(* IEC 61131-3 sources: Enumium/projects/downhome-spice-line/software/plc, 4 files *)

(* ---- DosingStation.st ---- *)
(* ============================================================================
   P1-225  PHASE 1 DOSING STATION  (IEC 61131-3 ST, CODESYS 3.5 on WAGO PFC200 750-8212)
   Down Home Creole Phase 1 prototype. Ring of up to 12 ingredient bins
   (P1-211) with 2 in volumetric screw feeders (P1-212, VFD P1-226) dosing
   one at a time into weigh hopper P1-220 (3 x 50 kg cells, Rice Lake 880
   indicator P1-222, 10 g division). When the list is done, butterfly valve
   P1-223 opens and flexible screw P1-224 carries the charge to blender P1-301
   (on riser stand P1-311). The hand-weighed lines and the premix are then
   tipped into the screw's intake grate, so nobody lifts a pail above waist height.

   The MES owns the recipe and the lot genealogy:
     GET /api/batch/<id>/doselist  -> MES_DoseList (largest dose first)
     POST /api/dose {batch, bin, actual_kg} after each finished dose.
   The PLC owns the equipment: one feeder at a time, never a screw into a
   closed valve or a full blender, no dose from a bin at low level.

   Dosing method (gain in weight, per bin):
     FAST  : VFD at FastHz until  net >= target - SlowBand - InFlight
     SLOW  : VFD at SlowHz until  net >= target - InFlight
     SETTLE: feeder off, wait SettleT, read stable weight
     CHECK : |actual - target| <= TolKg  -> report;  under -> one JOG pulse
             (max 3) ;  over -> OVERDOSE alarm, hold for the operator.
   In-flight (material still falling after the screw stops) is learned per
   bin: InFlight := InFlight + 0.5 * (actual - target), clamped 0..0.5 kg.
   No-flow: hopper gain < 0.05 kg in NoFlowT while the feeder runs -> alarm
   (bridged bin, empty bin, broken shear pin).
   Timers and speeds marked (SAT) are tuned at site acceptance.
   E-stop and the hopper/screw guards are hard-wired through safety relay
   SR-P1 and remove VFD enable; this code only sees the healthy bit.
   ============================================================================ *)

TYPE E_DoseStep : (
    IDLE := 0, WAIT_LIST := 5, PRECHECK := 10, TARE := 20, FAST := 30, SLOW := 40,
    SETTLE := 50, CHECK := 60, JOG := 65, REPORT := 70, NEXT := 80,
    TRANSFER := 90, TRANSFER_DRAIN := 95, COMPLETE := 100, HELD := 110, ABORTED := 120 );
END_TYPE

TYPE ST_DoseStep :
STRUCT
    Bin        : INT;          (* 1..12, ring position *)
    Ingredient : STRING[24];
    TargetKg   : REAL;         (* >= 4 kg by MES rule *)
    TolKg      : REAL;         (* max(1 % of target, 0.02 kg) *)
END_STRUCT
END_TYPE

TYPE ST_DoseList :
STRUCT
    BatchID  : STRING[16];
    FormulaID: STRING[16];
    Steps    : ARRAY[1..12] OF ST_DoseStep;
    Count    : INT;
    Valid    : BOOL;
END_STRUCT
END_TYPE

TYPE ST_DoseResult :
STRUCT
    BatchID  : STRING[16];
    Bin      : INT;
    ActualKg : REAL;
    Ready    : BOOL;           (* MES gateway posts /api/dose then sets Ack *)
    Ack      : BOOL;
END_STRUCT
END_TYPE

VAR_GLOBAL CONSTANT
    NBINS        : INT  := 12;
    HOPPER_MAXKG : REAL := 100.0;   (* 3 x 50 kg cells, 2/3 derated for the hopper *)
    BLENDER_MAXKG: REAL := 95.0;    (* P1-301 6 cu ft x densest blend (0.56 g/ml) *)
END_VAR

VAR_GLOBAL
    (* ---- I/O (WAGO 750-8212 rack: 750-430 DI, 750-530 DO, 750-455 AI 4-20 mA, Modbus RTU to GS20 drives) ---- *)
    DI_SafetyOK      AT %IX0.0  : BOOL;     (* SR-P1 healthy: e-stops, hopper lid, screw guard *)
    DI_ValveClosed   AT %IX0.1  : BOOL;     (* P1-223 closed limit *)
    DI_ValveOpen     AT %IX0.2  : BOOL;     (* P1-223 open limit *)
    DI_ScrewRunning  AT %IX0.3  : BOOL;     (* P1-224 motor contactor aux *)
    DI_BlenderReady  AT %IX0.4  : BOOL;     (* P1-301 cover closed and not discharging *)
    DI_BlenderHigh   AT %IX0.5  : BOOL;     (* P1-301 high level, capacitance probe *)
    DI_DustFanOn     AT %IX0.6  : BOOL;     (* P1-310 fan running *)
    DI_BinLow        AT %IX1.0  : ARRAY[1..12] OF BOOL;   (* P1-213 Soliphant FTM20, TRUE = covered (fail-safe) *)
    DO_ValveOpen     AT %QX0.0  : BOOL;     (* P1-223 solenoid *)
    DO_ScrewRun      AT %QX0.1  : BOOL;     (* P1-224 contactor *)
    DO_Horn          AT %QX0.2  : BOOL;
    DO_Beacon        AT %QX0.3  : BOOL;
    DO_Agitator      AT %QX1.0  : ARRAY[1..12] OF BOOL;   (* bin flow aid, density < 0.5 kg/L bins only *)
    AI_HopperKg                 : REAL;     (* P1-222 Rice Lake 880 gross weight over Modbus TCP, 10 g *)
    AI_HopperStable             : BOOL;     (* 880 motion bit inverted *)
    VFD_Run          : ARRAY[1..12] OF BOOL;      (* GS20 drives, Modbus RTU *)
    VFD_Hz           : ARRAY[1..12] OF REAL;
    VFD_Fault        : ARRAY[1..12] OF BOOL;

    (* ---- MES interface (OPC UA server on the PFC200, written by the MES gateway) ---- *)
    MES_DoseList     : ST_DoseList;
    MES_Result       : ST_DoseResult;
    MES_Start        : BOOL;
    MES_HandAddsDone : BOOL;            (* hand-weighed lines, then the premix, tipped into the P1-224 intake grate *)
    MES_Abort        : BOOL;
    HMI_Resume       : BOOL;
    HMI_Reset        : BOOL;

    (* ---- status ---- *)
    Dose_Step        : E_DoseStep;
    Dose_Index       : INT;
    Dose_NetKg       : REAL;
    Dose_Alarm       : STRING[60];
    Dose_HeldFrom    : E_DoseStep;

    (* ---- per-bin parameters, retained (learned in-flight survives power loss) ---- *)
    InFlightKg       : ARRAY[1..12] OF REAL := [12(0.15)];   (* (SAT) start value *)
    FastHz           : ARRAY[1..12] OF REAL := [12(60.0)];   (* about 700 L/h at 60 Hz, 2 in screw *)
    SlowHz           : ARRAY[1..12] OF REAL := [12(12.0)];   (* (SAT) *)
    SlowBandKg       : ARRAY[1..12] OF REAL := [12(1.0)];    (* (SAT) *)
END_VAR

PROGRAM DosingStation
VAR
    tStep     : TON;
    tNoFlow   : TON;
    tSettle   : TON;
    tTransfer : TON;
    TareKg    : REAL;
    LastKg    : REAL;
    ActualKg  : REAL;
    Jogs      : INT;
    i         : INT;
    b         : INT;           (* bin of the current step *)
    s         : ST_DoseStep;
    SumKg     : REAL;
    NoFlowT   : TIME := T#8S;  (* (SAT) *)
    SettleT   : TIME := T#3S;  (* (SAT) *)
    JogT      : TIME := T#600MS;
    DrainT    : TIME := T#20S; (* screw runs on after the hopper reads empty *)
    MaxDoseT  : TIME := T#10M; (* longest planned dose < 8 min *)
END_VAR

(* ---------- always: interlocks ---------- *)
IF NOT DI_SafetyOK OR MES_Abort THEN
    FOR i := 1 TO NBINS DO VFD_Run[i] := FALSE; END_FOR
    DO_ScrewRun := FALSE;
    DO_ValveOpen := FALSE;
    IF Dose_Step <> IDLE AND Dose_Step <> COMPLETE THEN
        Dose_Alarm := SEL(MES_Abort, 'SAFETY CIRCUIT OPEN', 'ABORTED BY MES');
        Dose_Step := ABORTED;
    END_IF
END_IF

(* the transfer screw may only run with the valve open, the blender ready and the dust fan on *)
IF DO_ScrewRun AND NOT (DI_ValveOpen AND DI_BlenderReady AND DI_DustFanOn AND NOT DI_BlenderHigh) THEN
    DO_ScrewRun := FALSE;
    DO_ValveOpen := FALSE;
    Dose_Alarm := 'TRANSFER PERMISSIVE LOST';
    Dose_HeldFrom := Dose_Step;
    Dose_Step := HELD;
END_IF

(* one feeder at a time: only the current bin may run *)
FOR i := 1 TO NBINS DO
    IF VFD_Run[i] AND ((Dose_Step <> FAST AND Dose_Step <> SLOW AND Dose_Step <> JOG) OR i <> b) THEN
        VFD_Run[i] := FALSE;
    END_IF
    IF VFD_Fault[i] AND VFD_Run[i] THEN
        VFD_Run[i] := FALSE;
        Dose_Alarm := CONCAT('FEEDER FAULT BIN ', INT_TO_STRING(i));
        Dose_HeldFrom := Dose_Step;
        Dose_Step := HELD;
    END_IF
    DO_Agitator[i] := VFD_Run[i];       (* flow aid only while its feeder runs *)
END_FOR

Dose_NetKg := AI_HopperKg - TareKg;

(* ---------- sequence ---------- *)
CASE Dose_Step OF

IDLE:
    IF MES_Start THEN Dose_Step := WAIT_LIST; END_IF

WAIT_LIST:
    IF MES_DoseList.Valid AND MES_DoseList.Count >= 1 AND MES_DoseList.Count <= NBINS THEN
        SumKg := 0.0;
        FOR i := 1 TO MES_DoseList.Count DO SumKg := SumKg + MES_DoseList.Steps[i].TargetKg; END_FOR
        IF SumKg > HOPPER_MAXKG OR SumKg > BLENDER_MAXKG THEN
            Dose_Alarm := 'DOSE LIST EXCEEDS HOPPER OR BLENDER';
            Dose_Step := ABORTED;
        ELSE
            Dose_Index := 1;
            Dose_Step := PRECHECK;
        END_IF
    END_IF

PRECHECK:
    (* hopper empty, valve closed, dust fan on *)
    IF NOT DI_DustFanOn THEN
        Dose_Alarm := 'DUST COLLECTOR P1-310 OFF';
    ELSIF NOT DI_ValveClosed THEN
        Dose_Alarm := 'HOPPER VALVE NOT CLOSED';
    ELSIF AI_HopperKg > 0.5 THEN
        Dose_Alarm := 'HOPPER NOT EMPTY';
    ELSE
        Dose_Alarm := '';
        Dose_Step := TARE;
    END_IF

TARE:
    s := MES_DoseList.Steps[Dose_Index];
    b := s.Bin;
    IF b < 1 OR b > NBINS THEN
        Dose_Alarm := 'BAD BIN NUMBER IN DOSE LIST';
        Dose_Step := ABORTED;
    ELSIF NOT DI_BinLow[b] THEN
        Dose_Alarm := CONCAT('BIN LOW: REFILL BIN ', INT_TO_STRING(b));   (* MES checked book stock; this is the probe *)
        Dose_HeldFrom := TARE;
        Dose_Step := HELD;
    ELSIF AI_HopperStable THEN
        TareKg := AI_HopperKg;        (* cumulative: each dose is tared on the previous ones *)
        LastKg := AI_HopperKg;
        Jogs := 0;
        VFD_Hz[b] := FastHz[b];
        VFD_Run[b] := TRUE;
        Dose_Step := FAST;
    END_IF

FAST, SLOW:
    IF Dose_Step = FAST AND Dose_NetKg >= s.TargetKg - SlowBandKg[b] - InFlightKg[b] THEN
        VFD_Hz[b] := SlowHz[b];
        Dose_Step := SLOW;
    ELSIF Dose_NetKg >= s.TargetKg - InFlightKg[b] THEN
        VFD_Run[b] := FALSE;
        Dose_Step := SETTLE;
    END_IF
    (* no-flow: the hopper must gain 50 g in NoFlowT *)
    tNoFlow(IN := VFD_Run[b] AND (AI_HopperKg - LastKg) < 0.05, PT := NoFlowT);
    IF (AI_HopperKg - LastKg) >= 0.05 THEN LastKg := AI_HopperKg; END_IF
    IF tNoFlow.Q THEN
        VFD_Run[b] := FALSE;
        Dose_Alarm := CONCAT('NO FLOW BIN ', INT_TO_STRING(b));
        Dose_HeldFrom := SLOW;    (* resume keeps TareKg and finishes the dose at slow speed *)
        Dose_Step := HELD;
    END_IF
    tStep(IN := TRUE, PT := MaxDoseT);
    IF tStep.Q THEN
        VFD_Run[b] := FALSE;
        Dose_Alarm := CONCAT('DOSE TIMEOUT BIN ', INT_TO_STRING(b));
        Dose_HeldFrom := SETTLE;
        Dose_Step := HELD;
    END_IF

SETTLE:
    tSettle(IN := AI_HopperStable, PT := SettleT);
    IF tSettle.Q THEN
        tSettle(IN := FALSE);
        ActualKg := AI_HopperKg - TareKg;
        Dose_Step := CHECK;
    END_IF

CHECK:
    IF ABS(ActualKg - s.TargetKg) <= s.TolKg THEN
        IF Jogs = 0 THEN
            (* learn in-flight only from clean single-shot doses *)
            InFlightKg[b] := LIMIT(0.0, InFlightKg[b] + 0.5 * (ActualKg - s.TargetKg), 0.5);
        END_IF
        Dose_Step := REPORT;
    ELSIF ActualKg < s.TargetKg - s.TolKg AND Jogs < 3 THEN
        Jogs := Jogs + 1;
        VFD_Hz[b] := SlowHz[b];
        VFD_Run[b] := TRUE;
        Dose_Step := JOG;
    ELSE
        (* over-dose or still short after 3 jogs: the operator corrects by hand at the hopper
           (scoop out or hand add on the 880) and resumes; the MES rejects anything outside tolerance *)
        Dose_Alarm := SEL(ActualKg > s.TargetKg, CONCAT('UNDERDOSE BIN ', INT_TO_STRING(b)), CONCAT('OVERDOSE BIN ', INT_TO_STRING(b)));
        Dose_HeldFrom := SETTLE;
        Dose_Step := HELD;
    END_IF

JOG:
    tStep(IN := TRUE, PT := JogT);
    IF tStep.Q THEN
        VFD_Run[b] := FALSE;
        Dose_Step := SETTLE;
    END_IF

REPORT:
    MES_Result.BatchID := MES_DoseList.BatchID;
    MES_Result.Bin := b;
    MES_Result.ActualKg := ActualKg;
    MES_Result.Ready := TRUE;
    IF MES_Result.Ack THEN
        MES_Result.Ready := FALSE;
        MES_Result.Ack := FALSE;
        Dose_Step := NEXT;
    END_IF

NEXT:
    IF Dose_Index < MES_DoseList.Count THEN
        Dose_Index := Dose_Index + 1;
        Dose_Step := TARE;
    ELSIF DI_BlenderReady AND NOT DI_BlenderHigh THEN
        DO_ValveOpen := TRUE;
        Dose_Step := TRANSFER;
    END_IF

TRANSFER:
    (* the bin charge goes first; the screw keeps running for the hand adds *)
    IF DI_ValveOpen THEN DO_ScrewRun := TRUE; END_IF
    IF AI_HopperKg < 0.2 AND AI_HopperStable THEN
        DO_ValveOpen := FALSE;
        Dose_Step := TRANSFER_DRAIN;
    END_IF

TRANSFER_DRAIN:
    (* operator tips the hand-weighed pails, then the premix last, into the P1-224 intake grate and
       confirms on the MES; the screw then runs on DrainT to empty the tube into the blender *)
    IF MES_HandAddsDone THEN
        tTransfer(IN := TRUE, PT := DrainT);
        IF tTransfer.Q THEN
            tTransfer(IN := FALSE);
            DO_ScrewRun := FALSE;
            MES_HandAddsDone := FALSE;
            Dose_Step := COMPLETE;
        END_IF
    END_IF

COMPLETE:
    MES_Start := FALSE;
    MES_DoseList.Valid := FALSE;
    IF HMI_Reset THEN Dose_Step := IDLE; Dose_Alarm := ''; END_IF

HELD:
    FOR i := 1 TO NBINS DO VFD_Run[i] := FALSE; END_FOR
    DO_ScrewRun := FALSE;
    IF HMI_Resume AND DI_SafetyOK THEN
        HMI_Resume := FALSE;
        Dose_Alarm := '';
        IF Dose_HeldFrom = SETTLE THEN
            Dose_Step := SETTLE;          (* re-weigh after the operator's correction *)
        ELSIF Dose_HeldFrom = TARE THEN
            Dose_Step := TARE;
        ELSIF Dose_HeldFrom = FAST OR Dose_HeldFrom = SLOW THEN
            LastKg := AI_HopperKg;
            VFD_Hz[b] := SlowHz[b];
            VFD_Run[b] := TRUE;
            Dose_Step := SLOW;
        ELSIF Dose_HeldFrom = TRANSFER THEN
            DO_ValveOpen := TRUE;
            Dose_Step := TRANSFER;
        ELSE
            Dose_Step := Dose_HeldFrom;
        END_IF
    END_IF

ABORTED:
    FOR i := 1 TO NBINS DO VFD_Run[i] := FALSE; END_FOR
    DO_ScrewRun := FALSE;
    DO_ValveOpen := FALSE;
    MES_Start := FALSE;
    IF HMI_Reset AND DI_SafetyOK THEN Dose_Step := IDLE; Dose_Alarm := ''; MES_Abort := FALSE; END_IF

END_CASE

(* step timers reset on every step change *)
IF Dose_Step <> FAST AND Dose_Step <> SLOW AND Dose_Step <> JOG THEN
    tStep(IN := FALSE);
    tNoFlow(IN := FALSE);
END_IF

DO_Beacon := Dose_Step = HELD OR Dose_Step = ABORTED;
DO_Horn := DO_Beacon AND NOT HMI_Reset;

(* ---- io_map.st ---- *)
(* Generated by gen_tags.py from design/io.json. Do not edit by hand. *)

VAR_GLOBAL (* PLC-601 physical I/O *)
    BD301_RUN              AT %IX1.0   : BOOL;  (* BD-301: bag dump screw running (aux contact); wire 601-01-00 *)
    BB302_RUN              AT %IX1.1   : BOOL;  (* BB-302: salt discharger screw running (aux contact); wire 601-01-01 *)
    SC304_RUN              AT %IX1.2   : BOOL;  (* SC-304: sifter motor running (aux contact); wire 601-01-02 *)
    FC307_RUN              AT %IX1.3   : BOOL;  (* FC-307: bag filler screw running (aux contact); wire 601-01-03 *)
    DC310_RUN              AT %IX1.4   : BOOL;  (* DC-310: dust collector fan running (aux contact); wire 601-01-04 *)
    BD301_LIDCLOSED        AT %IX1.5   : BOOL;  (* BD-301: bag dump grate lid closed; wire 601-01-05 *)
    BD301_DCFAN_RUN        AT %IX1.6   : BOOL;  (* BD-301: bag dump integral collector fan running; wire 601-01-06 *)
    BB302_SPOUT_CLOSED     AT %IX1.7   : BOOL;  (* BB-302: salt bag spout access door closed; wire 601-01-07 *)
    BB302_HOPPER_LOW       AT %IX1.8   : BOOL;  (* BB-302: salt outlet hopper low level; wire 601-01-08 *)
    RB303_RUN              AT %IX1.9   : BOOL;  (* RB-303: ribbon blender motor running; wire 601-01-09 *)
    RB303_COVER_CLOSED     AT %IX1.10  : BOOL;  (* RB-303: blender cover interlock closed (status; safety via SR-607); wire 601-01-10 *)
    RB303_VALVE_OPEN       AT %IX1.11  : BOOL;  (* RB-303: discharge valve open limit switch; wire 601-01-11 *)
    RB303_VALVE_CLOSED     AT %IX1.12  : BOOL;  (* RB-303: discharge valve closed limit switch; wire 601-01-12 *)
    SC304_OVERS_FULL       AT %IX1.13  : BOOL;  (* SC-304: sifter oversize bin full; wire 601-01-13 *)
    MD305_DETECT           AT %IX1.14  : BOOL;  (* MD-305: metal detected (reject cycle); wire 601-01-14 *)
    MD305_FAULT            AT %IX1.15  : BOOL;  (* MD-305: metal detector fault / not ready; wire 601-01-15 *)
    MD305_REJ_VERIFY       AT %IX2.0   : BOOL;  (* MD-305: reject valve reached reject position; wire 601-02-00 *)
    MD305_REJBIN_FULL      AT %IX2.1   : BOOL;  (* MD-305: locked reject container full; wire 601-02-01 *)
    FC307_HOPPER_HIGH      AT %IX2.2   : BOOL;  (* FC-307: screw inlet hopper high level; wire 601-02-02 *)
    FC307_HOPPER_LOW       AT %IX2.3   : BOOL;  (* FC-307: screw inlet hopper low level; wire 601-02-03 *)
    BF306_BAG_PRESENT      AT %IX2.4   : BOOL;  (* BF-306: bulk bag spout clamped / bag present; wire 601-02-04 *)
    BF306_FILL_DONE        AT %IX2.5   : BOOL;  (* BF-306: bag at target weight (from filler controller); wire 601-02-05 *)
    DC310_VENT_BURST       AT %IX2.6   : BOOL;  (* DC-310: explosion vent burst indicator; wire 601-02-06 *)
    DC310_ISO_CLOSED       AT %IX2.7   : BOOL;  (* DC-310: inlet isolation flap valve closed; wire 601-02-07 *)
    AC311_LOWPRESS         AT %IX2.8   : BOOL;  (* AC-311: plant air low pressure switch; wire 601-02-08 *)
    SR601_OK               AT %IX2.9   : BOOL;  (* SR-607: blending safety relay outputs on (all e-stops reset); wire 601-02-09 *)
    PB601_RESET            AT %IX2.10  : BOOL;  (* SR-607: safety reset push button (blue); wire 601-02-10 *)
    BD301_START            AT %QX4.0   : BOOL;  (* BD-301: bag dump screw start command; wire 601-04-00 *)
    BB302_START            AT %QX4.1   : BOOL;  (* BB-302: salt discharger screw start command; wire 601-04-01 *)
    SC304_START            AT %QX4.2   : BOOL;  (* SC-304: sifter motor start command; wire 601-04-02 *)
    FC307_START            AT %QX4.3   : BOOL;  (* FC-307: bag filler screw start command; wire 601-04-03 *)
    DC310_START            AT %QX4.4   : BOOL;  (* DC-310: dust collector fan start command; wire 601-04-04 *)
    RB303_START            AT %QX4.5   : BOOL;  (* RB-303: ribbon blender motor start; wire 601-04-05 *)
    RB303_VALVE_OPEN_SOL   AT %QX4.6   : BOOL;  (* RB-303: discharge valve open solenoid; wire 601-04-06 *)
    RB303_VALVE_CLOSE_SOL  AT %QX4.7   : BOOL;  (* RB-303: discharge valve close solenoid; wire 601-04-07 *)
    BF306_FILL_START       AT %QX4.8   : BOOL;  (* BF-306: start bag fill; wire 601-04-08 *)
    BF306_SEAL_INFLATE     AT %QX4.9   : BOOL;  (* BF-306: inflatable spout seal; wire 601-04-09 *)
    BF306_DENSIFY          AT %QX4.10  : BOOL;  (* BF-306: vibratory densification deck; wire 601-04-10 *)
    SL601_RED              AT %QX4.11  : BOOL;  (* CP-300: blending stack light red; wire 601-04-11 *)
    SL601_AMBER            AT %QX4.12  : BOOL;  (* CP-300: blending stack light amber; wire 601-04-12 *)
    SL601_GREEN            AT %QX4.13  : BOOL;  (* CP-300: blending stack light green; wire 601-04-13 *)
    SL601_HORN             AT %QX4.14  : BOOL;  (* CP-300: blending stack light horn; wire 601-04-14 *)
    RB303_WEIGHT           AT %IW6.0   : REAL;  (* RB-303: blender load cells 4-20 mA (lb); wire 601-06-00 *)
    RB303_AMPS             AT %IW6.1   : REAL;  (* RB-303: blender motor current 4-20 mA; wire 601-06-01 *)
    DC310_DP               AT %IW6.2   : REAL;  (* DC-310: filter differential pressure 4-20 mA (in w.c.); wire 601-06-02 *)
    AC311_PRESS            AT %IW6.3   : REAL;  (* AC-311: plant air header pressure 4-20 mA (psi); wire 601-06-03 *)
END_VAR

VAR_GLOBAL (* PLC-602 physical I/O *)
    BU401_RUN              AT %IX1.0   : BOOL;  (* BU-401: line A bag discharger screw running; wire 602-01-00 *)
    UN402_RUN              AT %IX1.1   : BOOL;  (* UN-402: unscrambler running; wire 602-01-01 *)
    BU502_RUN              AT %IX1.2   : BOOL;  (* BU-502: station B bag discharger screw running; wire 602-01-02 *)
    FL403_HOPPER_HIGH      AT %IX1.3   : BOOL;  (* FL-403: filler hopper high level; wire 602-01-03 *)
    FL403_HOPPER_LOW       AT %IX1.4   : BOOL;  (* FL-403: filler hopper low level; wire 602-01-04 *)
    NW501_HOPPER_HIGH      AT %IX1.5   : BOOL;  (* NW-501: station B hopper high level; wire 602-01-05 *)
    NW501_HOPPER_LOW       AT %IX1.6   : BOOL;  (* NW-501: station B hopper low level; wire 602-01-06 *)
    CV417_FAULT            AT %IX1.7   : BOOL;  (* CV-417: conveyor drive fault (any of 4); wire 602-01-07 *)
    FL403_READY            AT %IX1.8   : BOOL;  (* FL-403: FL-403 ready / running (OEM machine handshake); wire 602-01-08 *)
    FL403_FAULT            AT %IX1.9   : BOOL;  (* FL-403: FL-403 fault; wire 602-01-09 *)
    CP404_READY            AT %IX1.10  : BOOL;  (* CP-404: CP-404 ready / running (OEM machine handshake); wire 602-01-10 *)
    CP404_FAULT            AT %IX1.11  : BOOL;  (* CP-404: CP-404 fault; wire 602-01-11 *)
    IS405_READY            AT %IX1.12  : BOOL;  (* IS-405: IS-405 ready / running (OEM machine handshake); wire 602-01-12 *)
    IS405_FAULT            AT %IX1.13  : BOOL;  (* IS-405: IS-405 fault; wire 602-01-13 *)
    LB406_READY            AT %IX1.14  : BOOL;  (* LB-406: LB-406 ready / running (OEM machine handshake); wire 602-01-14 *)
    LB406_FAULT            AT %IX1.15  : BOOL;  (* LB-406: LB-406 fault; wire 602-01-15 *)
    CW409_READY            AT %IX2.0   : BOOL;  (* CW-409: CW-409 ready / running (OEM machine handshake); wire 602-02-00 *)
    CW409_FAULT            AT %IX2.1   : BOOL;  (* CW-409: CW-409 fault; wire 602-02-01 *)
    CE411_READY            AT %IX2.2   : BOOL;  (* CE-411: CE-411 ready / running (OEM machine handshake); wire 602-02-02 *)
    CE411_FAULT            AT %IX2.3   : BOOL;  (* CE-411: CE-411 fault; wire 602-02-03 *)
    CK412_READY            AT %IX2.4   : BOOL;  (* CK-412: CK-412 ready / running (OEM machine handshake); wire 602-02-04 *)
    CK412_FAULT            AT %IX2.5   : BOOL;  (* CK-412: CK-412 fault; wire 602-02-05 *)
    CS413_READY            AT %IX2.6   : BOOL;  (* CS-413: CS-413 ready / running (OEM machine handshake); wire 602-02-06 *)
    CS413_FAULT            AT %IX2.7   : BOOL;  (* CS-413: CS-413 fault; wire 602-02-07 *)
    PA414_READY            AT %IX2.8   : BOOL;  (* PA-414: PA-414 ready / running (OEM machine handshake); wire 602-02-08 *)
    PA414_FAULT            AT %IX2.9   : BOOL;  (* PA-414: PA-414 fault; wire 602-02-09 *)
    PL415_READY            AT %IX2.10  : BOOL;  (* PL-415: PL-415 ready / running (OEM machine handshake); wire 602-02-10 *)
    PL415_FAULT            AT %IX2.11  : BOOL;  (* PL-415: PL-415 fault; wire 602-02-11 *)
    NW501_READY            AT %IX2.12  : BOOL;  (* NW-501: NW-501 ready / running (OEM machine handshake); wire 602-02-12 *)
    NW501_FAULT            AT %IX2.13  : BOOL;  (* NW-501: NW-501 fault; wire 602-02-13 *)
    PE401_BLOCKED          AT %IX2.14  : BOOL;  (* CV-417: container present at filler infeed; wire 602-02-14 *)
    PE402_BLOCKED          AT %IX2.15  : BOOL;  (* CV-417: backup before capper; wire 602-02-15 *)
    PE403_BLOCKED          AT %IX3.0   : BOOL;  (* CV-417: backup before labeler; wire 602-03-00 *)
    PE404_BLOCKED          AT %IX3.1   : BOOL;  (* CV-417: label sensor confirm after labeler; wire 602-03-01 *)
    PE405_BLOCKED          AT %IX3.2   : BOOL;  (* CV-417: vision trigger; wire 602-03-02 *)
    PE406_BLOCKED          AT %IX3.3   : BOOL;  (* CV-417: reject confirm after vision reject; wire 602-03-03 *)
    PE407_BLOCKED          AT %IX3.4   : BOOL;  (* CV-417: checkweigher infeed spacing; wire 602-03-04 *)
    PE408_BLOCKED          AT %IX3.5   : BOOL;  (* CV-417: accumulation table full; wire 602-03-05 *)
    PE409_BLOCKED          AT %IX3.6   : BOOL;  (* CV-417: accumulation table low; wire 602-03-06 *)
    PE410_BLOCKED          AT %IX3.7   : BOOL;  (* CV-417: case infeed to sealer; wire 602-03-07 *)
    PE501_BLOCKED          AT %IX3.8   : BOOL;  (* NW-501: pouch at sealer infeed; wire 602-03-08 *)
    PE502_BLOCKED          AT %IX3.9   : BOOL;  (* NW-501: pouch out of sealer; wire 602-03-09 *)
    PE503_BLOCKED          AT %IX3.10  : BOOL;  (* NW-501: tub at fill station; wire 602-03-10 *)
    PE504_BLOCKED          AT %IX3.11  : BOOL;  (* NW-501: carton at fill station; wire 602-03-11 *)
    VS408_FAIL             AT %IX3.12  : BOOL;  (* VS-408: vision inspection fail; wire 602-03-12 *)
    CW409_BIN_FULL         AT %IX3.13  : BOOL;  (* CW-409: checkweigher locking reject bin full; wire 602-03-13 *)
    CW409_BIN_DOOR         AT %IX3.14  : BOOL;  (* CW-409: reject bin door closed and locked; wire 602-03-14 *)
    TT407_FAULT            AT %IX3.15  : BOOL;  (* TT-407: TTO coder fault / ribbon low; wire 602-03-15 *)
    TJ505_FAULT            AT %IX4.0   : BOOL;  (* TJ-505: TIJ coder fault / cartridge low; wire 602-04-00 *)
    SR602_OK               AT %IX4.1   : BOOL;  (* SR-607: line safety relay outputs on; wire 602-04-01 *)
    PB602_RESET            AT %IX4.2   : BOOL;  (* SR-607: safety reset push button (blue); wire 602-04-02 *)
    BU401_START            AT %QX5.0   : BOOL;  (* BU-401: line A bag discharger screw start; wire 602-05-00 *)
    UN402_START            AT %QX5.1   : BOOL;  (* UN-402: unscrambler start; wire 602-05-01 *)
    BU502_START            AT %QX5.2   : BOOL;  (* BU-502: station B bag discharger screw start; wire 602-05-02 *)
    CV417_RUN_CMD          AT %QX5.3   : BOOL;  (* CV-417: line A conveyor drives run; wire 602-05-03 *)
    FL403_PERMIT           AT %QX5.4   : BOOL;  (* FL-403: line permissive to FL-403; wire 602-05-04 *)
    CP404_PERMIT           AT %QX5.5   : BOOL;  (* CP-404: line permissive to CP-404; wire 602-05-05 *)
    IS405_PERMIT           AT %QX5.6   : BOOL;  (* IS-405: line permissive to IS-405; wire 602-05-06 *)
    LB406_PERMIT           AT %QX5.7   : BOOL;  (* LB-406: line permissive to LB-406; wire 602-05-07 *)
    CW409_PERMIT           AT %QX5.8   : BOOL;  (* CW-409: line permissive to CW-409; wire 602-05-08 *)
    CE411_PERMIT           AT %QX5.9   : BOOL;  (* CE-411: line permissive to CE-411; wire 602-05-09 *)
    CK412_PERMIT           AT %QX5.10  : BOOL;  (* CK-412: line permissive to CK-412; wire 602-05-10 *)
    CS413_PERMIT           AT %QX5.11  : BOOL;  (* CS-413: line permissive to CS-413; wire 602-05-11 *)
    PA414_PERMIT           AT %QX5.12  : BOOL;  (* PA-414: line permissive to PA-414; wire 602-05-12 *)
    PL415_PERMIT           AT %QX5.13  : BOOL;  (* PL-415: line permissive to PL-415; wire 602-05-13 *)
    NW501_PERMIT           AT %QX5.14  : BOOL;  (* NW-501: line permissive to NW-501; wire 602-05-14 *)
    RJ408_FIRE             AT %QX5.15  : BOOL;  (* VS-408: reject pusher after vision; wire 602-05-15 *)
    SL602_RED              AT %QX6.0   : BOOL;  (* CP-400: line A stack light red; wire 602-06-00 *)
    SL602_AMBER            AT %QX6.1   : BOOL;  (* CP-400: line A stack light amber; wire 602-06-01 *)
    SL602_GREEN            AT %QX6.2   : BOOL;  (* CP-400: line A stack light green; wire 602-06-02 *)
    SL602_HORN             AT %QX6.3   : BOOL;  (* CP-400: line A stack light horn; wire 602-06-03 *)
END_VAR

(* ---- BlendTrain.st ---- *)
(* ============================================================================
   PLC-601  BLENDING TRAIN SEQUENCE  (ISA-88 phase logic, IEC 61131-3 ST)
   Down Home Creole dry plant. Train: BD-301 / BB-302 -> RB-303 -> SC-304 ->
   DH-102 magnet -> MD-305 (CCP-1) -> FC-307 -> BF-306.
   Tags come from io_map.st (generated from design/io.json).

   The MES (software/mes) owns the recipe. It downloads one batch at a time:
   BatchID, FormulaID, TargetKg, MixTime_s, SaltKg, AllergenClass. The PLC
   owns equipment safety: it will not open a cover, run a screw into a closed
   valve, or fill a bag that MD-305 has not cleared.
   ============================================================================ *)

TYPE E_BlendStep : (
    IDLE := 0, WAIT_DOWNLOAD := 5, PRECHECK := 10, CHARGE_SALT := 20,
    CHARGE_MAJORS := 30, CHARGE_PREMIX := 40, MIX := 50, HOLD_SAMPLE := 55,
    DISCHARGE := 60, DRAIN := 70, PURGE := 80, COMPLETE := 90,
    HELD := 100, ABORTED := 110 );
END_TYPE

TYPE ST_BatchDownload :
STRUCT
    BatchID       : STRING[16];   (* DHyyjjj-B## *)
    FormulaID     : STRING[16];
    TargetKg      : REAL;         (* <= RB-303 working volume x bulk density, checked by MES and here *)
    SaltKg        : REAL;         (* metered by BB-302 on blender load cells *)
    MixTime_s     : DINT;         (* site: 12 min *)
    AllergenClass : INT;          (* 0 none, 1 wheat (Friday campaign only) *)
    Valid         : BOOL;
END_STRUCT
END_TYPE

VAR_GLOBAL
    MES_Download    : ST_BatchDownload;   (* written by MES over OPC UA / CIP *)
    MES_MajorsDone  : BOOL;               (* operator scanned all major bags at BD-301 *)
    MES_PremixDone  : BOOL;               (* premix bag scanned and dumped *)
    MES_SampleOK    : BOOL;               (* QC accepted in-process sample (optional hold) *)
    MES_Abort       : BOOL;
    Blend_Step      : E_BlendStep;
    Blend_StateText : STRING[40];
    Blend_ActKg     : REAL;
    Blend_SaltActKg : REAL;
    Blend_MixLeft_s : DINT;
    Blend_Alarm     : WORD;               (* bit map, see ALARMS below *)
    MD305_RejCount  : DINT;               (* reported to MES for the batch record *)
    BlendMaxKg      : REAL := 655.0;      (* 36 cu ft working (1,019 L) x 0.643 g/mL densest formula; MES checks the formula-specific limit first *)
END_VAR

PROGRAM BlendTrain
VAR
    tMix        : TON;
    tDrain      : TON;
    tPurge      : TON;
    tValve      : TON;
    tamps       : TON;
    WeightAtStart : REAL;
    Permissive  : BOOL;
    DustOK      : BOOL;
    rDetect     : R_TRIG;
    rReset      : R_TRIG;
END_VAR

(* ---------- PERMISSIVES (hard interlocks also exist in safety relay SR-601) ---------- *)
DustOK := DC310_RUN AND NOT DC310_ISO_CLOSED (* flap valve trips closed on deflagration *) AND NOT DC310_VENT_BURST AND DC310_DP > 0.5 AND DC310_DP < 6.0;  (* in. w.c. *)
Permissive := SR601_OK AND DustOK AND NOT AC311_LOWPRESS AND RB303_COVER_CLOSED AND NOT MD305_FAULT;

(* Weight from RB-303 load cells (AI, kg) *)
Blend_ActKg := RB303_WEIGHT;

(* ---------- ALARMS ---------- *)
Blend_Alarm.0 := NOT SR601_OK;           (* e-stop / guard *)
Blend_Alarm.1 := NOT DustOK;             (* dust collector not proven or vent burst: NFPA 652 *)
Blend_Alarm.2 := AC311_LOWPRESS;
Blend_Alarm.3 := NOT RB303_COVER_CLOSED;
Blend_Alarm.4 := MD305_FAULT;
Blend_Alarm.5 := MD305_REJBIN_FULL;
Blend_Alarm.6 := SC304_OVERS_FULL;
Blend_Alarm.7 := BB302_HOPPER_LOW AND Blend_Step = CHARGE_SALT;
Blend_Alarm.8 := tamps.Q;                (* blender over-current: possible lump or overfill *)
tamps(IN := RB303_AMPS > 24.0, PT := T#5S);  (* M-304 FLA 21 A *)

rReset(CLK := PB601_RESET);
rDetect(CLK := MD305_DETECT);
IF rDetect.Q THEN MD305_RejCount := MD305_RejCount + 1; END_IF;

(* Any loss of permissive while running -> HELD with every mover stopped *)
IF NOT Permissive AND Blend_Step > PRECHECK AND Blend_Step < COMPLETE THEN
    Blend_Step := HELD;
END_IF;
IF MES_Abort AND Blend_Step <> IDLE THEN
    Blend_Step := ABORTED;
END_IF;

CASE Blend_Step OF
IDLE:
    Blend_StateText := 'Idle';
    IF MES_Download.Valid THEN Blend_Step := PRECHECK; END_IF;

PRECHECK:
    Blend_StateText := 'Pre-check';
    (* batch size never above blender working capacity (design-basis batch rule) *)
    IF MES_Download.TargetKg > BlendMaxKg OR MES_Download.TargetKg <= 0.0 THEN
        Blend_Alarm.9 := TRUE; MES_Download.Valid := FALSE; Blend_Step := IDLE;
    ELSIF Permissive AND RB303_VALVE_CLOSED AND Blend_ActKg < 5.0 THEN
        WeightAtStart := Blend_ActKg; MD305_RejCount := 0;
        Blend_Step := CHARGE_SALT;
    END_IF;

CHARGE_SALT:
    Blend_StateText := 'Charging salt (BB-302)';
    RB303_START := TRUE;                    (* ribbons turn during charge to avoid salt bed *)
    BB302_START := (Blend_ActKg - WeightAtStart) < (MES_Download.SaltKg - 3.0);  (* 3 kg in-flight, tuned at SAT *)
    IF NOT BB302_START THEN
        Blend_SaltActKg := Blend_ActKg - WeightAtStart;
        Blend_Step := CHARGE_MAJORS;
    END_IF;

CHARGE_MAJORS:
    Blend_StateText := 'Dump majors at BD-301';
    BD301_START := BD301_DCFAN_RUN;  (* screw runs only with the station dust fan proven *)
    IF MES_MajorsDone THEN BD301_START := FALSE; Blend_Step := CHARGE_PREMIX; END_IF;

CHARGE_PREMIX:
    Blend_StateText := 'Add premix at BD-301';
    BD301_START := BD301_DCFAN_RUN;
    IF MES_PremixDone THEN
        BD301_START := FALSE;
        tMix(IN := FALSE);
        Blend_Step := MIX;
    END_IF;

MIX:
    Blend_StateText := 'Mixing';
    RB303_START := TRUE;
    tMix(IN := TRUE, PT := DINT_TO_TIME(MES_Download.MixTime_s * 1000));
    Blend_MixLeft_s := MES_Download.MixTime_s - TIME_TO_DINT(tMix.ET) / 1000;
    IF tMix.Q THEN tMix(IN := FALSE); Blend_Step := HOLD_SAMPLE; END_IF;

HOLD_SAMPLE:
    Blend_StateText := 'Sample for CV (QC)';
    RB303_START := FALSE;
    IF MES_SampleOK THEN Blend_Step := DISCHARGE; END_IF;

DISCHARGE:
    Blend_StateText := 'Discharging to bulk bag';
    (* start downstream first, then open valve: no product into a stopped screw *)
    IF NOT BF306_BAG_PRESENT THEN
        Blend_Alarm.10 := TRUE;
    ELSE
        Blend_Alarm.10 := FALSE;
        BF306_SEAL_INFLATE := TRUE;
        FC307_START := NOT FC307_HOPPER_LOW OR SC304_RUN;
        SC304_START := TRUE;
        RB303_START := TRUE;
        BF306_DENSIFY := TRUE;
        BF306_FILL_START := TRUE;
        (* throttle: close blender valve while FC-307 hopper is high *)
        RB303_VALVE_OPEN_SOL := SC304_RUN AND FC307_RUN AND NOT FC307_HOPPER_HIGH AND NOT MD305_REJBIN_FULL;
        RB303_VALVE_CLOSE_SOL := NOT RB303_VALVE_OPEN_SOL;
        tValve(IN := RB303_VALVE_OPEN_SOL AND NOT RB303_VALVE_OPEN, PT := T#3S);
        Blend_Alarm.11 := tValve.Q;   (* valve did not prove open *)
        IF Blend_ActKg < 2.0 THEN tDrain(IN := FALSE); Blend_Step := DRAIN; END_IF;
    END_IF;

DRAIN:
    Blend_StateText := 'Draining train';
    RB303_VALVE_OPEN_SOL := FALSE; RB303_VALVE_CLOSE_SOL := TRUE;
    tDrain(IN := TRUE, PT := T#90S);      (* sifter and screw run empty *)
    IF tDrain.Q THEN
        SC304_START := FALSE; FC307_START := FALSE; RB303_START := FALSE;
        BF306_FILL_START := FALSE; BF306_DENSIFY := FALSE;
        tDrain(IN := FALSE); Blend_Step := COMPLETE;
    END_IF;

COMPLETE:
    Blend_StateText := 'Complete: release bag to HOLD-1';
    BF306_SEAL_INFLATE := NOT BF306_FILL_DONE;
    MES_Download.Valid := FALSE; MES_MajorsDone := FALSE; MES_PremixDone := FALSE; MES_SampleOK := FALSE;
    Blend_Step := IDLE;

HELD:
    Blend_StateText := 'HELD: check alarms, press reset';
    BD301_START := FALSE; BB302_START := FALSE; SC304_START := FALSE; FC307_START := FALSE;
    RB303_START := FALSE; RB303_VALVE_OPEN_SOL := FALSE; RB303_VALVE_CLOSE_SOL := TRUE;
    BF306_FILL_START := FALSE; BF306_DENSIFY := FALSE;
    (* resume at charge step if material was already weighed; MES knows which step *)
    IF rReset.Q AND Permissive THEN Blend_Step := MIX; END_IF;

ABORTED:
    Blend_StateText := 'ABORTED: batch on hold in MES';
    BD301_START := FALSE; BB302_START := FALSE; SC304_START := FALSE; FC307_START := FALSE;
    RB303_START := FALSE; RB303_VALVE_OPEN_SOL := FALSE; RB303_VALVE_CLOSE_SOL := TRUE;
    BF306_FILL_START := FALSE;
    IF rReset.Q THEN MES_Abort := FALSE; MES_Download.Valid := FALSE; Blend_Step := IDLE; END_IF;
END_CASE;

(* Dust collector always runs while any mover runs, and 10 min after (post-purge) *)
DC310_START := SR601_OK AND NOT DC310_VENT_BURST AND (Blend_Step <> IDLE OR BD301_DCFAN_RUN);

(* Stack light *)
SL601_RED   := Blend_Alarm <> 0 OR Blend_Step = HELD OR Blend_Step = ABORTED;
SL601_AMBER := Blend_Step = CHARGE_MAJORS OR Blend_Step = CHARGE_PREMIX OR Blend_Step = HOLD_SAMPLE;
SL601_GREEN := Blend_Step = MIX OR Blend_Step = DISCHARGE OR Blend_Step = DRAIN;
SL601_HORN  := Blend_Alarm.1 OR Blend_Alarm.5;   (* dust and reject-bin full sound locally *)
END_PROGRAM

(* ---- PackLineA.st ---- *)
(* ============================================================================
   PLC-602  PACK LINE A  -  PackML (ISA-TR88.00.02) state machine + line control
   BU-401 > FL-403 > CP-404 > IS-405 > LB-406/TT-407 > VS-408/RJ-408 > CW-409 >
   AT-410 > CE-411/CK-412 > CS-413 > PA-414 > PL-415
   Each OEM machine keeps its own controller and guarding. This PLC gives each
   one a PERMIT and reads READY/FAULT, runs the conveyor, the vision reject and
   the backup/starve logic, and exchanges the job with the MES.
   ============================================================================ *)

TYPE E_PackML : (
    STOPPED := 2, STARTING := 3, IDLE := 4, SUSPENDED := 5, EXECUTE := 6,
    STOPPING := 7, ABORTING := 8, ABORTED := 9, HOLDING := 10, HELD := 11,
    UNHOLDING := 12, SUSPENDING := 13, UNSUSPENDING := 14, RESETTING := 15,
    COMPLETING := 16, COMPLETE := 17, CLEARING := 1 );
END_TYPE

TYPE ST_Job :
STRUCT
    JobID        : STRING[20];
    SKU          : STRING[16];
    LotCode      : STRING[24];    (* DHyyjjj-B## + BEST BY text sent to TT-407 *)
    BlendBagID   : STRING[20];    (* released FIBC; BU-401 scan must match *)
    Container    : INT;           (* 1 shaker-250, 2 shaker-320, 3 jar-12 ... selects change-part recipe *)
    NetG         : REAL;
    TargetG      : REAL;          (* net x (1 + overfill) *)
    TareG        : REAL;
    UnitsOrdered : DINT;
    CaseCount    : INT;
    SpeedUPM     : REAL;          (* 80 shakers / 45 jars, from line balance *)
    Valid        : BOOL;
END_STRUCT
END_TYPE

VAR_GLOBAL
    MES_Job         : ST_Job;
    MES_BagScanOK   : BOOL;         (* MES confirms FIBC at BU-401 is released and matches job *)
    MES_LabelOK     : BOOL;         (* MES confirms first-off label/lot code check signed *)
    Cmd_Start, Cmd_Stop, Cmd_Reset, Cmd_Hold, Cmd_Unhold, Cmd_Abort, Cmd_Clear : BOOL;
    LineA_State     : E_PackML := STOPPED;
    LineA_Good      : DINT;         (* accepted by CW-409 *)
    LineA_RejVision : DINT;
    LineA_RejWeight : DINT;         (* counted by CW-409 over OPC UA, mirrored here *)
    LineA_Cases     : DINT;
    LineA_StopReason: INT;          (* first-out, for OEE in MES *)
    LineA_MachSpeed : REAL;         (* upm command to FL-403 *)
END_VAR

PROGRAM PackLineA
VAR
    Faults      : WORD;
    AllReady    : BOOL;
    Starved     : BOOL;
    Blocked     : BOOL;
    tStarve     : TON;
    tBlock      : TON;
    tStep       : TON;
    tRejChk     : TON;      (* reject must be confirmed by PE-406 within 500 ms *)
    rVis        : R_TRIG;
    rCase       : R_TRIG;
    rReset      : R_TRIG;
    RejQueue    : ARRAY[0..15] OF BOOL;   (* shift register: vision fail -> pusher, 6 pitches *)
    rPitch      : R_TRIG;
    i           : INT;
END_VAR

(* ---------- machine status ---------- *)
Faults.0  := FL403_FAULT;  Faults.1 := CP404_FAULT;  Faults.2 := IS405_FAULT;  Faults.3 := LB406_FAULT;
Faults.4  := CW409_FAULT;  Faults.5 := CE411_FAULT;  Faults.6 := CK412_FAULT;  Faults.7 := CS413_FAULT;
Faults.8  := PA414_FAULT;  Faults.9 := PL415_FAULT;  Faults.10 := CV417_FAULT; Faults.11 := TT407_FAULT;
Faults.12 := CW409_BIN_FULL OR CW409_BIN_DOOR;   (* reject bin must be locked and not full: CCP verification *)
Faults.13 := NOT SR602_OK;
Faults.14 := tRejChk.Q;   (* pusher fired but PE-406 did not see the reject *)

AllReady := FL403_READY AND CP404_READY AND IS405_READY AND LB406_READY AND CW409_READY
            AND CE411_READY AND CK412_READY AND CS413_READY AND PA414_READY AND PL415_READY;

(* first-out stop reason *)
IF LineA_StopReason = 0 AND Faults <> 0 THEN
    FOR i := 0 TO 15 DO
        IF (WORD_TO_DINT(SHR(Faults, i)) MOD 2) = 1 AND LineA_StopReason = 0 THEN LineA_StopReason := i + 1; END_IF;
    END_FOR;
END_IF;

(* starve: filler hopper low with no bag running; block: accumulation full *)
tStarve(IN := FL403_HOPPER_LOW AND NOT BU401_RUN, PT := T#20S);   Starved := tStarve.Q;
tBlock(IN := PE408_BLOCKED, PT := T#5S);                           Blocked := tBlock.Q;

rReset(CLK := Cmd_Reset OR PB602_RESET);

(* ---------- global transitions ---------- *)
IF Faults.13 OR Cmd_Abort THEN
    IF LineA_State <> ABORTED THEN LineA_State := ABORTING; END_IF;
ELSIF Faults <> 0 AND (LineA_State = EXECUTE OR LineA_State = SUSPENDED OR LineA_State = STARTING) THEN
    LineA_State := HOLDING;
ELSIF Cmd_Stop AND LineA_State <> STOPPED AND LineA_State <> ABORTED THEN
    LineA_State := STOPPING;
END_IF;

CASE LineA_State OF
STOPPED:
    IF rReset.Q THEN LineA_State := RESETTING; END_IF;

RESETTING:
    LineA_StopReason := 0;
    IF AllReady AND SR602_OK THEN LineA_State := IDLE; END_IF;

IDLE:
    (* job, released bag and signed first-off label are all required before start *)
    IF Cmd_Start AND MES_Job.Valid AND MES_BagScanOK AND MES_LabelOK THEN
        tStep(IN := FALSE); LineA_State := STARTING;
    END_IF;

STARTING:
    CV417_RUN_CMD := TRUE;
    tStep(IN := TRUE, PT := T#3S);           (* conveyor first, then machines, downstream to upstream *)
    IF tStep.Q THEN tStep(IN := FALSE); LineA_State := EXECUTE; END_IF;

EXECUTE:
    LineA_MachSpeed := MES_Job.SpeedUPM;
    IF Starved OR Blocked THEN LineA_State := SUSPENDING; END_IF;
    IF LineA_Good >= MES_Job.UnitsOrdered THEN LineA_State := COMPLETING; END_IF;

SUSPENDING:  LineA_State := SUSPENDED;
SUSPENDED:
    LineA_MachSpeed := 0.0;
    IF NOT Starved AND NOT Blocked THEN LineA_State := UNSUSPENDING; END_IF;
UNSUSPENDING: LineA_State := EXECUTE;

HOLDING:     LineA_State := HELD;
HELD:
    IF Faults = 0 AND (Cmd_Unhold OR rReset.Q) THEN LineA_State := UNHOLDING; END_IF;
UNHOLDING:   LineA_State := EXECUTE;

COMPLETING:
    (* run out: stop filler, keep downstream running until accumulation empties *)
    LineA_MachSpeed := 0.0;
    tStep(IN := NOT PE409_BLOCKED, PT := T#30S);
    IF tStep.Q THEN tStep(IN := FALSE); LineA_State := COMPLETE; END_IF;
COMPLETE:
    MES_Job.Valid := FALSE; MES_BagScanOK := FALSE; MES_LabelOK := FALSE;
    IF rReset.Q THEN LineA_State := RESETTING; END_IF;

STOPPING:    LineA_MachSpeed := 0.0; LineA_State := STOPPED;
ABORTING:    LineA_MachSpeed := 0.0; LineA_State := ABORTED;
ABORTED:
    IF Cmd_Clear AND SR602_OK THEN LineA_State := CLEARING; END_IF;
CLEARING:    LineA_State := STOPPED;
END_CASE;

(* ---------- outputs ---------- *)
CV417_RUN_CMD := LineA_State = STARTING OR LineA_State = EXECUTE OR LineA_State = SUSPENDED
                 OR LineA_State = COMPLETING OR LineA_State = UNSUSPENDING OR LineA_State = UNHOLDING;
FL403_PERMIT  := LineA_State = EXECUTE AND NOT PE402_BLOCKED;      (* no fill into a backed-up capper *)
BU401_START   := (LineA_State = EXECUTE OR LineA_State = SUSPENDED) AND MES_BagScanOK AND NOT FL403_HOPPER_HIGH;
UN402_START   := LineA_State = EXECUTE AND NOT PE401_BLOCKED;
CP404_PERMIT  := CV417_RUN_CMD;
IS405_PERMIT  := CV417_RUN_CMD;
LB406_PERMIT  := CV417_RUN_CMD AND NOT TT407_FAULT;                 (* never label without a lot code *)
CW409_PERMIT  := CV417_RUN_CMD;
CE411_PERMIT  := CV417_RUN_CMD;
CK412_PERMIT  := CV417_RUN_CMD;
CS413_PERMIT  := CV417_RUN_CMD;
PA414_PERMIT  := CV417_RUN_CMD;
PL415_PERMIT  := LineA_State <> ABORTED AND SR602_OK;

(* vision reject: shift register clocked by vision trigger eye, pusher 6 pitches downstream *)
rVis(CLK := PE405_BLOCKED);
IF rVis.Q THEN
    FOR i := 15 TO 1 BY -1 DO RejQueue[i] := RejQueue[i - 1]; END_FOR;
    RejQueue[0] := VS408_FAIL;
    IF VS408_FAIL THEN LineA_RejVision := LineA_RejVision + 1; END_IF;
END_IF;
RJ408_FIRE := RejQueue[6] AND PE405_BLOCKED;
tRejChk(IN := (RJ408_FIRE OR tRejChk.IN) AND NOT PE406_BLOCKED, PT := T#500MS);

rCase(CLK := PE410_BLOCKED);
IF rCase.Q THEN LineA_Cases := LineA_Cases + 1; END_IF;

SL602_RED   := LineA_State = HELD OR LineA_State = ABORTED OR LineA_State = STOPPED;
SL602_AMBER := LineA_State = SUSPENDED OR LineA_State = IDLE OR LineA_State = COMPLETE;
SL602_GREEN := LineA_State = EXECUTE;
SL602_HORN  := LineA_State = ABORTING OR Faults.12;
END_PROGRAM
